// TIA Portal V20 export
DATA_BLOCK "06_Grundstellungen_DB"   // DB177
// stored: InstanceOfName 06_Grundstellungen, InstanceOfType FB
"06_Grundstellungen"
BEGIN
END_DATA_BLOCK
